(*
SPDX-FileCopyrightText: c 2026 Oleksandr Tiutyk <trofimich@gmail.com>
SPDX-License-Identifier: MIT
License: https://opensource.org/license/mit
*)

(*!
<summary>Checks generic membership with independent borrowed queries.</summary>
<description>
Borrows a group-owned stack reserved for this case. Use from one task at a stable address.
Teardown clears the stack and test-owned resources before publication.
</description>
*)

{attribute 'no_assign'}
{attribute 'no_explicit_call' := 'do not call this function block directly'}
FUNCTION_BLOCK StackContainsGenericTest EXTENDS TOF_Testing.SingleCycleTest
VAR_STAT
	{attribute 'hide'}
	_ClassName : STRING := __POUNAME();
END_VAR
VAR
	_Stack : TOF_Collections.IStack;
END_VAR

(*!
<summary>Clears the fixture before the runner publishes the result.</summary>
<description>
Also runs after an unexpected exception interrupts the case.
</description>
*)
METHOD PROTECTED AfterTest
_Stack.Clear();
END_METHOD

//! <summary>Borrows the concrete class name. Callers must not modify it.</summary>
{attribute 'monitoring' := 'call'}
PROPERTY ClassName : REFERENCE TO STRING
GET
ClassName REF= _ClassName;
END_GET
END_PROPERTY

(*!
<summary>Checks generic membership with independent borrowed queries.</summary>
*)
METHOD PROTECTED ExecuteTest
VAR
	values : ARRAY [1..4] OF INT := [11, 22, 33, 44];
	query : TOF_Core.GENERIC_VALUE;
END_VAR
_Stack.PushCopy(value := values[1]);
_Stack.PushCopy(value := values[2]);
_Stack.PushCopy(value := values[3]);

query := TOF_Core.GenericValueFactory.FromIntReference(value := values[1]);
Assert.ThatBool(
	actual := _Stack.ContainsGeneric(value := query, releaseValue := FALSE),
	message := "Generic lookup must find the bottom value"
).IsTrue();

query := TOF_Core.GenericValueFactory.FromIntReference(value := values[3]);
Assert.ThatBool(
	actual := _Stack.ContainsGeneric(value := query, releaseValue := FALSE),
	message := "Generic lookup must find the top value"
).IsTrue();

query := TOF_Core.GenericValueFactory.FromIntReference(value := values[4]);
Assert.ThatBool(
	actual := _Stack.ContainsGeneric(value := query, releaseValue := FALSE),
	message := "Generic lookup must reject an absent value"
).IsFalse();

Assert.ThatDInt(
	actual := _Stack.Length,
	message := "Generic lookup must preserve all three entries"
).ToBe(expected := DINT#3);
END_METHOD

(*!
<summary>Binds the stack fixture for this case.</summary>
<description>
Stores a borrowed interface without invoking the fixture. The owning group keeps it alive and
reserves it for this case. TestElement initializes the name and parent.
</description>
<param name="name">Display name of this case.</param>
<param name="parent">Group that owns this case.</param>
<param name="stack">Required live stack reserved for this case.</param>
*)
METHOD FB_init : BOOL
VAR_INPUT
	bInitRetains: BOOL; // TRUE: the retain variables are initialized (reset warm / reset cold)
	bInCopyCode: BOOL; // TRUE: the instance will be copied to the copy code afterward (online change)
	name : WSTRING;
	parent : TOF_Testing.ITestElement;
	stack : TOF_Collections.IStack;
END_VAR
_Stack := stack;
FB_init := TRUE;
END_METHOD

//! <summary>Borrows the compiler-initialized namespace name. Callers must not modify it.</summary>
{attribute 'monitoring' := 'call'}
PROPERTY NamespaceName : REFERENCE TO STRING
GET
NamespaceName REF= CurrentNamespace.Name;
END_GET
END_PROPERTY

//! <summary>Reports the concrete instance size in bytes.</summary>
{attribute 'monitoring' := 'call'}
PROPERTY SelfSize : ULINT
GET
SelfSize := XSIZEOF(THIS^);
END_GET
END_PROPERTY

END_FUNCTION_BLOCK

(* stored: Version 1.1.0.1, ProductVersion 3.1.4026.21
   POU StackContainsGenericTest: Id {e62e0d15-4c09-4c6f-8464-ee19a383eb4a}, SpecialFunc None
   Method AfterTest: Id {284d2fbd-3145-432f-8c4a-c129d33b8eca}
   Property ClassName: Id {8836ae1b-67aa-4b7c-9f04-dfec30089881}
   Get Get: Id {60e96e51-6ae7-4680-a8cb-7b457511a340}
   Method ExecuteTest: Id {6c147a1e-b27b-4cbb-a0d2-4099e4ca71ef}
   Method FB_init: Id {4d63b32f-2dcd-42ab-ba61-089d2d63aa22}
   Property NamespaceName: Id {38c2e328-3cac-4969-839f-13b7b925bf16}
   Get Get: Id {c5c70f06-ac4f-4814-9d8a-718176a0cea3}
   Property SelfSize: Id {5b6497b0-b6e0-494f-80bf-0136aad47c65}
   Get Get: Id {4cf4eb27-0d43-4057-9f97-addfb307de1d} *)
